(* IEC 61131-3 sources: kns-pump-station/src/GVLs/Station, 2 files *)

(* ---- GVL_Station.gvl.st ---- *)
// Назначение: данные обмена станции с HMI, OPC UA и MQTT (04 §19.1). Команды пишут клиенты,
//             остальное пишет только PRG_Station.
// Автор:      kr0nsch
// Версия:     0.1.0
// Документ:   docs/DESIGN.md, раздел 4.1
{attribute 'qualified_only'}
VAR_GLOBAL
    stStationCmd    : ST_StationCmd;     // команды (ReadWrite в символах)
    stStationSts    : ST_StationSts;     // состояние (Read)
    fbLIC101        : PL.FB_PID;         // регулятор уровня; HMI и SCADA читают fbLIC101.stSts
    stLIC101Cmd     : PL.ST_PidCmd;      // команды фейсплейта LIC101 (ReadWrite)
    fbAlarms        : FB_StationAlarms;  // тревоги KNS1.* (источник для сводки)
    // диагностика для HMI и OPC UA (пишет только PRG_Station)
    axPumpRun       : ARRAY[1..GVL_Const.STN_PUMP_COUNT] OF BOOL;   // → fbP10n.xAutoRun
    awPumpInterlock : ARRAY[1..GVL_Const.STN_PUMP_COUNT] OF WORD;   // → fbP10n.wInterlock
    rSpeedSp_pct    : REAL;                                         // → fbP10n.rSpeedSpAuto_pct
    stCfgLkg        : ST_StationCfg;     // последняя корректная копия уставок (Read)
END_VAR

(* ---- GVL_StationDefaults.gvl.st ---- *)
// Назначение: уставки станции и LIC101 по умолчанию — команда «Применить уставки проекта»
//             (GVL_Hmi.xApplyProjectCfg, 04 §18.3). Имена — как у переменных GVL_Persist; значения
//             LIC101 — тот же инициализатор, что в блоке станции GVL_Persist (DESIGN, раздел 4.7):
//             их совпадение сверяет тест StationDefaultsMatchPersistInit.
// Автор:      kr0nsch
// Версия:     0.1.0
// Документ:   docs/DESIGN.md, раздел 4.2
{attribute 'qualified_only'}
VAR_GLOBAL CONSTANT
    // Умолчания типа (раздел 3.1). Инициализатор нужен компилятору (без него C0228); остальные поля —
    // умолчания ST_StationCfg, совпадение с типом сверяет тест StationDefaultsMatchTypeDefaults.
    // lint:allow STL007 имя как у переменной GVL_Persist (DESIGN 4.2)
    stStationCfg : ST_StationCfg := (eRotation := E_RotationMode.RunHours);
    // lint:allow STL007 имя как у переменной GVL_Persist (DESIGN 4.2); LIC101 (04 §18.2, № 32–43)
    stLIC101Cfg  : PL.ST_PidCfg := (
        eAction := PL.E_PidAction.Direct, rKp := 6.0, rTi_s := 600.0, rTd_s := 0.0,
        rPvMin_eu := 0.0, rPvMax_eu := 5.0, rSpMin_eu := 1.2, rSpMax_eu := 2.2,
        rOutMin_pct := 0.0, rOutMax_pct := 100.0, tSample := T#500MS,
        ePvFailAction := PL.E_PidPvFailAction.Hold, rSafeOut_pct := 100.0, xUseOutAct := TRUE,
        udiAlarmIdBase := 100100,
        astAlarm := [(ePriority := PL.E_AlarmPriority.None), (ePriority := PL.E_AlarmPriority.None),
                     (ePriority := PL.E_AlarmPriority.None), (ePriority := PL.E_AlarmPriority.None),
                     (ePriority := PL.E_AlarmPriority.None), (ePriority := PL.E_AlarmPriority.None),
                     (ePriority := PL.E_AlarmPriority.None), (ePriority := PL.E_AlarmPriority.None)]);
END_VAR
